(* IEC 61131-3 sources: PLC-Static-Analysis/modules/plc-rules/src/test/resources/PLCA-Q002/strict, 1 file *)

(* ---- strict.st ---- *)
TYPE E_Light : (Red, Green); END_TYPE

PROGRAM P_Strict
VAR
    eLight : E_Light;
    b : BOOL;
END_VAR
CASE eLight OF // PLCA-Q002
    Red: b := FALSE;
    Green: b := TRUE;
END_CASE
END_PROGRAM
